(* IEC 61131-3 sources: plc-st-coding-agent/progress/evidence/f14_v11_public_20261113/jobs/codex_deepseek-v4pro, 8 files *)

(* ---- public-easy-01.candidate_01.st ---- *)
FUNCTION_BLOCK FillingLineControl
VAR_INPUT
    bottleSensor : BOOL;
    cleaningConfirmButton : BOOL;
    fillingConfirmButton : BOOL;
    cappingConfirmButton : BOOL;
    packingConfirmButton : BOOL;
    finishedButton : BOOL;
END_VAR
VAR_OUTPUT
    Pump_Motor : BOOL;
    Filling_Valve : BOOL;
    Capping_Machine : BOOL;
    Packing_Machine : BOOL;
    Completion_Light : BOOL;
END_VAR
VAR
    stage : INT := 0;
END_VAR

(*
ENGINEERING_CONTRACT
Output           Activation / Retention / Explicit Deactivation / Same-Scan Priority
Pump_Motor:      activ=stage0 + bottleSensor (PUB001); hold=stage1; deact=cleaningConfirm -> stage2 (PUB002).
Filling_Valve:   activ=cleaningConfirm at stage1 (PUB002); hold=stage2; deact=fillingConfirm -> stage3 (PUB003).
Capping_Machine: activ=fillingConfirm at stage2 (PUB003); hold=stage3; deact=cappingConfirm -> stage4 (PUB004).
Packing_Machine: activ=cappingConfirm at stage3 (PUB004); hold=stage4; deact=packingConfirm -> stage5 (PUB005).
Completion_Light: activ=packingConfirm at stage4 (PUB005); hold=stage5; deact=finishedButton -> stage0 (PUB006).
All states retained in local stage; outputs mutually exclusive. Same scan: finished reset evaluated first, then bottle and sequence transitions. No physical units/timers.
*)

(* CONTRACT_RULES [] *)

IF finishedButton AND (stage = 5) THEN
    stage := 0;
END_IF;

IF bottleSensor AND (stage = 0) THEN
    stage := 1;
END_IF;

IF cleaningConfirmButton AND (stage = 1) THEN
    stage := 2;
END_IF;

IF fillingConfirmButton AND (stage = 2) THEN
    stage := 3;
END_IF;

IF cappingConfirmButton AND (stage = 3) THEN
    stage := 4;
END_IF;

IF packingConfirmButton AND (stage = 4) THEN
    stage := 5;
END_IF;

Pump_Motor := (stage = 1);
Filling_Valve := (stage = 2);
Capping_Machine := (stage = 3);
Packing_Machine := (stage = 4);
Completion_Light := (stage = 5);

END_FUNCTION_BLOCK

(* ---- public-easy-01.candidate_02.st ---- *)
FUNCTION_BLOCK FillingLineControl
VAR_INPUT
    bottleSensor : BOOL;
    cleaningConfirmButton : BOOL;
    fillingConfirmButton : BOOL;
    cappingConfirmButton : BOOL;
    packingConfirmButton : BOOL;
    finishedButton : BOOL;
END_VAR
VAR_OUTPUT
    Pump_Motor : BOOL;
    Filling_Valve : BOOL;
    Capping_Machine : BOOL;
    Packing_Machine : BOOL;
    Completion_Light : BOOL;
END_VAR
VAR
    stage : INT := 0;
END_VAR

(*
ENGINEERING_CONTRACT
Output           Activation / Retention / Explicit Deactivation / Same-Scan Priority
Pump_Motor:      activ=stage0 + bottleSensor (PUB001); hold=stage1; deact=cleaningConfirm -> stage2 (PUB004).
Filling_Valve:   activ=cleaningConfirm at stage1 (PUB004); hold=stage2; deact=fillingConfirm -> stage3 (PUB003).
Capping_Machine: activ=fillingConfirm at stage2 (PUB003); hold=stage3; deact=cappingConfirm -> stage4 (PUB004).
Packing_Machine: activ=cappingConfirm at stage3 (PUB004); hold=stage4; deact=packingConfirm -> stage5 (PUB005).
Completion_Light: activ=packingConfirm at stage4 (PUB005); hold=stage5; deact=finishedButton -> stage0 (PUB006).
All states retained in local stage; outputs mutually exclusive. Same scan: finished reset evaluated first, then one eligible sequence transition is applied.
*)

(* CONTRACT_RULES [] *)

IF finishedButton AND (stage = 5) THEN
    stage := 0;
END_IF;

IF (stage = 0) AND bottleSensor THEN
    stage := 1;
ELSIF (stage = 1) AND cleaningConfirmButton THEN
    stage := 2;
ELSIF (stage = 2) AND fillingConfirmButton THEN
    stage := 3;
ELSIF (stage = 3) AND cappingConfirmButton THEN
    stage := 4;
ELSIF (stage = 4) AND packingConfirmButton THEN
    stage := 5;
END_IF;

Pump_Motor := (stage = 1);
Filling_Valve := (stage = 2);
Capping_Machine := (stage = 3);
Packing_Machine := (stage = 4);
Completion_Light := (stage = 5);

END_FUNCTION_BLOCK

(* ---- public-easy-01.raw_candidate_01.st ---- *)
FUNCTION_BLOCK FillingLineControl
VAR_INPUT
    bottleSensor : BOOL;
    cleaningConfirmButton : BOOL;
    fillingConfirmButton : BOOL;
    cappingConfirmButton : BOOL;
    packingConfirmButton : BOOL;
    finishedButton : BOOL;
END_VAR
VAR_OUTPUT
    Pump_Motor : BOOL;
    Filling_Valve : BOOL;
    Capping_Machine : BOOL;
    Packing_Machine : BOOL;
    Completion_Light : BOOL;
END_VAR
VAR
    stage : INT := 0;
END_VAR

(*
ENGINEERING_CONTRACT
Output           Activation / Retention / Explicit Deactivation / Same-Scan Priority
Pump_Motor:      activ=stage0 + bottleSensor (PUB001); hold=stage1; deact=cleaningConfirm -> stage2 (PUB002).
Filling_Valve:   activ=cleaningConfirm at stage1 (PUB002); hold=stage2; deact=fillingConfirm -> stage3 (PUB003).
Capping_Machine: activ=fillingConfirm at stage2 (PUB003); hold=stage3; deact=cappingConfirm -> stage4 (PUB004).
Packing_Machine: activ=cappingConfirm at stage3 (PUB004); hold=stage4; deact=packingConfirm -> stage5 (PUB005).
Completion_Light: activ=packingConfirm at stage4 (PUB005); hold=stage5; deact=finishedButton -> stage0 (PUB006).
All states retained in local stage; outputs mutually exclusive. Same scan: finished reset evaluated first, then bottle and sequence transitions. No physical units/timers.
*)

(* CONTRACT_RULES [] *)

IF finishedButton AND (stage = 5) THEN
    stage := 0;
END_IF;

IF bottleSensor AND (stage = 0) THEN
    stage := 1;
END_IF;

IF cleaningConfirmButton AND (stage = 1) THEN
    stage := 2;
END_IF;

IF fillingConfirmButton AND (stage = 2) THEN
    stage := 3;
END_IF;

IF cappingConfirmButton AND (stage = 3) THEN
    stage := 4;
END_IF;

IF packingConfirmButton AND (stage = 4) THEN
    stage := 5;
END_IF;

Pump_Motor := (stage = 1);
Filling_Valve := (stage = 2);
Capping_Machine := (stage = 3);
Packing_Machine := (stage = 4);
Completion_Light := (stage = 5);

END_FUNCTION_BLOCK

(* ---- public-easy-01.raw_candidate_02.st ---- *)
FUNCTION_BLOCK FillingLineControl
VAR_INPUT
    bottleSensor : BOOL;
    cleaningConfirmButton : BOOL;
    fillingConfirmButton : BOOL;
    cappingConfirmButton : BOOL;
    packingConfirmButton : BOOL;
    finishedButton : BOOL;
END_VAR
VAR_OUTPUT
    Pump_Motor : BOOL;
    Filling_Valve : BOOL;
    Capping_Machine : BOOL;
    Packing_Machine : BOOL;
    Completion_Light : BOOL;
END_VAR
VAR
    stage : INT := 0;
END_VAR

(*
ENGINEERING_CONTRACT
Output           Activation / Retention / Explicit Deactivation / Same-Scan Priority
Pump_Motor:      activ=stage0 + bottleSensor (PUB001); hold=stage1; deact=cleaningConfirm -> stage2 (PUB004).
Filling_Valve:   activ=cleaningConfirm at stage1 (PUB004); hold=stage2; deact=fillingConfirm -> stage3 (PUB003).
Capping_Machine: activ=fillingConfirm at stage2 (PUB003); hold=stage3; deact=cappingConfirm -> stage4 (PUB004).
Packing_Machine: activ=cappingConfirm at stage3 (PUB004); hold=stage4; deact=packingConfirm -> stage5 (PUB005).
Completion_Light: activ=packingConfirm at stage4 (PUB005); hold=stage5; deact=finishedButton -> stage0 (PUB006).
All states retained in local stage; outputs mutually exclusive. Same scan: finished reset evaluated first, then one eligible sequence transition is applied.
*)

(* CONTRACT_RULES [] *)

IF finishedButton AND (stage = 5) THEN
    stage := 0;
END_IF;

IF (stage = 0) AND bottleSensor THEN
    stage := 1;
ELSIF (stage = 1) AND cleaningConfirmButton THEN
    stage := 2;
ELSIF (stage = 2) AND fillingConfirmButton THEN
    stage := 3;
ELSIF (stage = 3) AND cappingConfirmButton THEN
    stage := 4;
ELSIF (stage = 4) AND packingConfirmButton THEN
    stage := 5;
END_IF;

Pump_Motor := (stage = 1);
Filling_Valve := (stage = 2);
Capping_Machine := (stage = 3);
Packing_Machine := (stage = 4);
Completion_Light := (stage = 5);

END_FUNCTION_BLOCK

(* ---- public-easy-02.candidate_01.st ---- *)
(* ENGINEERING_CONTRACT
   hasChanged: activation when current DWORD differs from stored previous scan; combinational, not held.
   hasRisingEdges/risingBits/noOfRisingBits: activation for 0->1 bits versus prior scan; computed each scan, not held.
   hasFallingEdges/fallingBits/noOfFallingBits: activation for 1->0 bits versus prior scan; computed each scan, not held.
   Retention/hold: only prevValue is retained; outputs are overwritten every scan from current comparison.
   Explicit reset/deactivation: none defined in PUB001; first scan establishes baseline with no edge/changed outputs.
   Same-scan priority: current value is compared against retained prior word before prior word is updated.
   Units/boundaries: DWORD bits 0..31, USINT counts 0..32, zero-based bit iteration.
*)
(* CONTRACT_RULES [] *)
FUNCTION_BLOCK FB
VAR
    prevValue : DWORD;
    isInitialized : BOOL;
    tmpRising : DWORD;
    tmpFalling : DWORD;
    tmpBitIndex : INT;
END_VAR

IF NOT isInitialized THEN
    hasChanged := FALSE;
    hasRisingEdges := FALSE;
    risingBits := DWORD#0;
    noOfRisingBits := 0;
    hasFallingEdges := FALSE;
    fallingBits := DWORD#0;
    noOfFallingBits := 0;
    prevValue := value;
    isInitialized := TRUE;
    RETURN;
END_IF;

hasChanged := value <> prevValue;
tmpRising := value AND (NOT prevValue);
tmpFalling := prevValue AND (NOT value);

risingBits := tmpRising;
fallingBits := tmpFalling;
hasRisingEdges := tmpRising <> DWORD#0;
hasFallingEdges := tmpFalling <> DWORD#0;

noOfRisingBits := 0;
noOfFallingBits := 0;

FOR tmpBitIndex := 0 TO 31 DO
    IF (tmpRising AND SHL(DWORD#1, TO_DINT(tmpBitIndex))) <> DWORD#0 THEN
        noOfRisingBits := TO_USINT(noOfRisingBits + 1);
    END_IF;
    IF (tmpFalling AND SHL(DWORD#1, TO_DINT(tmpBitIndex))) <> DWORD#0 THEN
        noOfFallingBits := TO_USINT(noOfFallingBits + 1);
    END_IF;
END_FOR;

prevValue := value;

END_FUNCTION_BLOCK

(* ---- public-easy-02.candidate_02.st ---- *)
(* ENGINEERING_CONTRACT
   hasChanged: activation when current DWORD differs from stored previous scan; combinational, not held.
   hasRisingEdges/risingBits/noOfRisingBits: activation for 0->1 bits versus prior scan; computed each scan, not held.
   hasFallingEdges/fallingBits/noOfFallingBits: activation for 1->0 bits versus prior scan; computed each scan, not held.
   Retention/hold: only prevValue is retained; outputs are overwritten every scan from current comparison.
   Explicit reset/deactivation: none defined in PUB001; first scan establishes baseline with no edge/changed outputs.
   Same-scan priority: current value is compared against retained prior word before prior word is updated.
   Units/boundaries: DWORD bits 0..31, USINT counts 0..32, zero-based bit iteration.
*)
(* CONTRACT_RULES [] *)
FUNCTION_BLOCK FB
VAR_INPUT
    value : DWORD;
END_VAR
VAR_OUTPUT
    hasChanged : BOOL;
    hasRisingEdges : BOOL;
    risingBits : DWORD;
    noOfRisingBits : USINT;
    hasFallingEdges : BOOL;
    fallingBits : DWORD;
    noOfFallingBits : USINT;
END_VAR
VAR
    prevValue : DWORD;
    isInitialized : BOOL;
    tmpRising : DWORD;
    tmpFalling : DWORD;
    tmpBitIndex : INT;
END_VAR

IF NOT isInitialized THEN
    hasChanged := FALSE;
    hasRisingEdges := FALSE;
    risingBits := DWORD#0;
    noOfRisingBits := 0;
    hasFallingEdges := FALSE;
    fallingBits := DWORD#0;
    noOfFallingBits := 0;
    prevValue := value;
    isInitialized := TRUE;
    RETURN;
END_IF;

hasChanged := value <> prevValue;
tmpRising := value AND (NOT prevValue);
tmpFalling := prevValue AND (NOT value);

risingBits := tmpRising;
fallingBits := tmpFalling;
hasRisingEdges := tmpRising <> DWORD#0;
hasFallingEdges := tmpFalling <> DWORD#0;

noOfRisingBits := 0;
noOfFallingBits := 0;

FOR tmpBitIndex := 0 TO 31 DO
    IF (tmpRising AND SHL(DWORD#1, TO_DINT(tmpBitIndex))) <> DWORD#0 THEN
        noOfRisingBits := TO_USINT(noOfRisingBits + 1);
    END_IF;
    IF (tmpFalling AND SHL(DWORD#1, TO_DINT(tmpBitIndex))) <> DWORD#0 THEN
        noOfFallingBits := TO_USINT(noOfFallingBits + 1);
    END_IF;
END_FOR;

prevValue := value;

END_FUNCTION_BLOCK

(* ---- public-easy-02.raw_candidate_01.st ---- *)
(* ENGINEERING_CONTRACT
   hasChanged: activation when current DWORD differs from stored previous scan; combinational, not held.
   hasRisingEdges/risingBits/noOfRisingBits: activation for 0->1 bits versus prior scan; computed each scan, not held.
   hasFallingEdges/fallingBits/noOfFallingBits: activation for 1->0 bits versus prior scan; computed each scan, not held.
   Retention/hold: only prevValue is retained; outputs are overwritten every scan from current comparison.
   Explicit reset/deactivation: none defined in PUB001; first scan establishes baseline with no edge/changed outputs.
   Same-scan priority: current value is compared against retained prior word before prior word is updated.
   Units/boundaries: DWORD bits 0..31, USINT counts 0..32, zero-based bit iteration.
*)
(* CONTRACT_RULES [] *)
FUNCTION_BLOCK FB
VAR
    prevValue : DWORD;
    isInitialized : BOOL;
    tmpRising : DWORD;
    tmpFalling : DWORD;
    tmpBitIndex : INT;
END_VAR

IF NOT isInitialized THEN
    hasChanged := FALSE;
    hasRisingEdges := FALSE;
    risingBits := DWORD#0;
    noOfRisingBits := 0;
    hasFallingEdges := FALSE;
    fallingBits := DWORD#0;
    noOfFallingBits := 0;
    prevValue := value;
    isInitialized := TRUE;
    RETURN;
END_IF;

hasChanged := value <> prevValue;
tmpRising := value AND (NOT prevValue);
tmpFalling := prevValue AND (NOT value);

risingBits := tmpRising;
fallingBits := tmpFalling;
hasRisingEdges := tmpRising <> DWORD#0;
hasFallingEdges := tmpFalling <> DWORD#0;

noOfRisingBits := 0;
noOfFallingBits := 0;

FOR tmpBitIndex := 0 TO 31 DO
    IF (tmpRising AND SHL(DWORD#1, TO_DINT(tmpBitIndex))) <> DWORD#0 THEN
        noOfRisingBits := TO_USINT(noOfRisingBits + 1);
    END_IF;
    IF (tmpFalling AND SHL(DWORD#1, TO_DINT(tmpBitIndex))) <> DWORD#0 THEN
        noOfFallingBits := TO_USINT(noOfFallingBits + 1);
    END_IF;
END_FOR;

prevValue := value;

END_FUNCTION_BLOCK

(* ---- public-easy-02.raw_candidate_02.st ---- *)
(* ENGINEERING_CONTRACT
   hasChanged: activation when current DWORD differs from stored previous scan; combinational, not held.
   hasRisingEdges/risingBits/noOfRisingBits: activation for 0->1 bits versus prior scan; computed each scan, not held.
   hasFallingEdges/fallingBits/noOfFallingBits: activation for 1->0 bits versus prior scan; computed each scan, not held.
   Retention/hold: only prevValue is retained; outputs are overwritten every scan from current comparison.
   Explicit reset/deactivation: none defined in PUB001; first scan establishes baseline with no edge/changed outputs.
   Same-scan priority: current value is compared against retained prior word before prior word is updated.
   Units/boundaries: DWORD bits 0..31, USINT counts 0..32, zero-based bit iteration.
*)
(* CONTRACT_RULES [] *)
FUNCTION_BLOCK FB
VAR_INPUT
    value : DWORD;
END_VAR
VAR_OUTPUT
    hasChanged : BOOL;
    hasRisingEdges : BOOL;
    risingBits : DWORD;
    noOfRisingBits : USINT;
    hasFallingEdges : BOOL;
    fallingBits : DWORD;
    noOfFallingBits : USINT;
END_VAR
VAR
    prevValue : DWORD;
    isInitialized : BOOL;
    tmpRising : DWORD;
    tmpFalling : DWORD;
    tmpBitIndex : INT;
END_VAR

IF NOT isInitialized THEN
    hasChanged := FALSE;
    hasRisingEdges := FALSE;
    risingBits := DWORD#0;
    noOfRisingBits := 0;
    hasFallingEdges := FALSE;
    fallingBits := DWORD#0;
    noOfFallingBits := 0;
    prevValue := value;
    isInitialized := TRUE;
    RETURN;
END_IF;

hasChanged := value <> prevValue;
tmpRising := value AND (NOT prevValue);
tmpFalling := prevValue AND (NOT value);

risingBits := tmpRising;
fallingBits := tmpFalling;
hasRisingEdges := tmpRising <> DWORD#0;
hasFallingEdges := tmpFalling <> DWORD#0;

noOfRisingBits := 0;
noOfFallingBits := 0;

FOR tmpBitIndex := 0 TO 31 DO
    IF (tmpRising AND SHL(DWORD#1, TO_DINT(tmpBitIndex))) <> DWORD#0 THEN
        noOfRisingBits := TO_USINT(noOfRisingBits + 1);
    END_IF;
    IF (tmpFalling AND SHL(DWORD#1, TO_DINT(tmpBitIndex))) <> DWORD#0 THEN
        noOfFallingBits := TO_USINT(noOfFallingBits + 1);
    END_IF;
END_FOR;

prevValue := value;

END_FUNCTION_BLOCK
